(* IEC 61131-3 sources: NachHouse_TST/API/pilot_Api_V11, 8 files *)

(* ---- 07_Nh_JsonRamTest.st ---- *)
// One-shot transport measurement. The records are synthetic because the production mRam is not populated yet.
// Files intentionally remain in //RAM/NACHHOUSE/ for manual inspection after the test.

TYPE
  NH_REC_ALL {PUBLIC}  {HIDDEN}: STRUCT 	// uvodny zaznam pre vsetky DEV alebo struktury, ktore su tabulkou
 	  Ok              : BOOL := TRUE; // platna veta = NOT DELTED
    ID              : INT;					// identifikator zaznamu {Rec Number}
  END_STRUCT;

  NH_CFG_ALL	{PUBLIC}  {HIDDEN}: STRUCT 	// univerzalne CFG pre vsetky DEV
    RoomID          : INT;			    // do ktorej miestnosti patri toto DEV
    CategoryID      : INT;					// domovska kategoria Device
  END_STRUCT;

  NH_JSON_TEST_ROOM  {PUBLIC} : STRUCT    // povodna testovacia struktura
    // povodna testovacia struktura
    RoomId          : UDINT;
    LightLevel      : UINT;
    Temperature10   : INT;
    Online          : BOOL;
   END_STRUCT

  NH_JSON_MEM  {PUBLIC} : STRUCT    // toto zoberiema ako STATE  a bude cele v mRam ako struktura, ktora sa bude posielat do JSON-stat
    rec             : NH_REC_ALL;   // hlavicka - ked sa bude posielat do JSON len stat = mRam
    all             : NH_CFG_ALL;   // premenn, ktore sa pouzivaju casto pri behu programu, ale nemenia sa
    sta             : NH_JSON_TEST_ROOM;   // hlavnme stavove premenne
   END_STRUCT

  NH_JSON_TEST_ROOM_CFG {PUBLIC} : STRUCT   // konfiguracia ulozena
    rec             : NH_REC_ALL;   // duplicitna hlavicka - ked sa bude posielat do JSON len config
    Name            : STRING[32];  // nazov miestnosti
    // iba pre testivanie  STRUCT <-> JSON (ostatnych elementarnych typov, ktore mozu byt STRUCT -> JSON)
    _Dint           : DINT;
    _Sint           : SINT;
    _Usint          : USINT;
    _Uint           : USINT;
    _Real           : REAL;
    _LReal          : LREAL;
    _String         : STRING[30];   // prazdny string
    _StringCZSK     : STRING := 'SVKBEGIN_ščľťžýáíé_SVKEND';   // string obsahujuci ceske a slovenske znaky
    _BYTE           : BYTE;
    _WORD           : WORD;
    _TIME           : TIME;
    _DATE           : DATE;
    _TIME_OF_DAY    : TOD;
    _DATE_AND_TIME  : DT;
   END_STRUCT

  NH_LIGT {PUBLIC}  : STRUCT    // toto je kompletna premenn v nasom pripade JSON, inak NH_ROOM, NH_BLIND,NH_HEAT ...
    mem             : NH_JSON_MEM;             // co budes v mRam ako STATE (memory) - RAM je pouzita na disku '/RAM/'
    cfg             : NH_JSON_TEST_ROOM_CFG;   // toto bude len na SDC
   END_STRUCT

(*
   NH_JSON_TEST_ROOM : STRUCT
      RoomId          : UDINT;
      LightLevel      : UINT;
      Temperature10   : INT;
      Online          : BOOL;
   END_STRUCT
*)
END_TYPE

VAR_GLOBAL CONSTANT
  NH_JSON_TEST_RECORDS : UINT := 300;
  // Historical prototype declaration; unused and not valid in VAR_GLOBAL CONSTANT.
  // aNhJSON {PUBLIC} {TRACK_ADR} {OPEN_UP} : NH_LIGHT;
END_VAR

VAR_GLOBAL
   NhJsonTestRooms        : ARRAY[1..300] OF NH_JSON_TEST_ROOM;
   NhJsonTestInitialized  : BOOL := FALSE;
   NhJsonTestState        : USINT := 0;
   NhJsonTestMode         : USINT := 0;
   NhJsonTestIndex        : UINT := 0;
   NhJsonTestHandle       : HANDLE := INVALID_HANDLE_VALUE;
   NhJsonTestWritten      : UDINT := 0;
   NhJsonTestBuildCycles  : UINT := 0;
   NhJsonTestFileName     : STRING[80];
END_VAR

FUNCTION NhJsonTestWrite : BOOL
   VAR_INPUT
      Text : STRING[255];
   END_VAR
   VAR
      Count : UDINT;
   END_VAR
   NhJsonTestWrite := FALSE;
   Count := FileWrite(hFile := NhJsonTestHandle, adrBuf := PTR_TO_UDINT(ADR(Text)), size := UINT_TO_UDINT(LEN(Text)));
   IF Count <> UINT_TO_UDINT(LEN(Text)) THEN RETURN; END_IF;
   NhJsonTestWritten := NhJsonTestWritten + Count;
   NhJsonTestWrite := TRUE;
END_FUNCTION

FUNCTION NhJsonTestWriteRecord : BOOL
   VAR_INPUT
      Index  : UINT;
      Prefix : BOOL;
   END_VAR
   VAR
      Record : PTR_TO NH_JSON_TEST_ROOM;
      Line   : STRING[255];
      Online : STRING[5];
   END_VAR
   NhJsonTestWriteRecord := FALSE;
   Record := ADR(NhJsonTestRooms[Index]);
   IF Record^.Online THEN Online := 'true'; ELSE Online := 'false'; END_IF;
   IF Prefix THEN Line := ','; ELSE Line := ''; END_IF;
   Line := CONCAT(Line, '{"id":', UDINT_TO_STRING(Record^.RoomId), ',"level":', UINT_TO_STRING(Record^.LightLevel), ',"temperature10":', INT_TO_STRING(Record^.Temperature10), ',"online":', Online, '}');
   NhJsonTestWriteRecord := NhJsonTestWrite(Text := Line);
END_FUNCTION

FUNCTION NhJsonTestInitialize : BOOL
   VAR
      Index : UINT;
   END_VAR
   NhJsonTestInitialize := NhJsonTestInitialized;
   IF NhJsonTestInitialized THEN RETURN; END_IF;
   FOR Index := 1 TO NH_JSON_TEST_RECORDS DO
      NhJsonTestRooms[Index].RoomId := UINT_TO_UDINT(Index);
      NhJsonTestRooms[Index].LightLevel := (Index * 7) MOD 101;
      NhJsonTestRooms[Index].Temperature10 := 185 + UINT_TO_INT(Index MOD 65);
      NhJsonTestRooms[Index].Online := (Index MOD 11) <> 0;
   END_FOR;
   NhJsonTestInitialized := TRUE;
   NhJsonTestInitialize := TRUE;
END_FUNCTION

FUNCTION NhJsonTestCycle : BOOL
   VAR
      Index : UINT;
      Header : STRING[255];
      Trailer : STRING[255];
      ModeText : STRING[6];
      Closed : BOOL;
   END_VAR
   NhJsonTestCycle := FALSE;
   NhJsonTestInitialize();
   IF System_S.LAST_CYCLE_TIME_100US > NhJsonTestMaxCycle100us THEN NhJsonTestMaxCycle100us := System_S.LAST_CYCLE_TIME_100US; END_IF;
   CASE NhJsonTestState OF
      0:
         IF (NhJsonTestCommand = 1) OR (NhJsonTestCommand = 2) THEN
            NhJsonTestMode := NhJsonTestCommand; NhJsonTestCommand := 0; NhJsonTestStatus := NhJsonTestMode;
            NhJsonTestBytes := 0; NhJsonTestRecords := 0; NhJsonTestMaxCycle100us := 0; NhJsonTestWritten := 0; NhJsonTestBuildCycles := 0; NhJsonTestState := 1;
         END_IF;
      1:
         IF NhJsonTestMode = 1 THEN NhJsonTestFileName := '//RAM/NACHHOUSE/nh-json-test-stream.json'; ELSE NhJsonTestFileName := '//RAM/NACHHOUSE/nh-json-test-burst.json'; END_IF;
         NhJsonTestHandle := FileOpen(fileName := NhJsonTestFileName, mode := F_WRITE);
         IF NhJsonTestHandle = INVALID_HANDLE_VALUE THEN NhJsonTestStatus := 255; NhJsonTestState := 0; RETURN; END_IF;
         IF NhJsonTestMode = 1 THEN
            ModeText := 'stream';
         ELSE
            ModeText := 'burst';
         END_IF;
         Header := CONCAT('{"protocol":1,"kind":"patch","sequence":', UDINT_TO_STRING(NhTxRevision + 1), ',"baseSequence":', UDINT_TO_STRING(NhTxRevision), ',"mode":"', ModeText, '","groups":[{"type":"ROOMS","schema":"NH_JSON_TEST_ROOM","records":[');
         IF NOT NhJsonTestWrite(Text := Header) THEN NhJsonTestStatus := 255; NhJsonTestState := 4; RETURN; END_IF;
         NhJsonTestIndex := 1; NhJsonTestState := 2;
      2:
         IF NhJsonTestMode = 1 THEN
            IF NOT NhJsonTestWriteRecord(Index := NhJsonTestIndex, Prefix := NhJsonTestIndex > 1) THEN NhJsonTestStatus := 255; NhJsonTestState := 4; RETURN; END_IF;
            NhJsonTestIndex := NhJsonTestIndex + 1; NhJsonTestBuildCycles := NhJsonTestBuildCycles + 1;
         ELSE
            FOR Index := 1 TO NH_JSON_TEST_RECORDS DO
               IF NOT NhJsonTestWriteRecord(Index := Index, Prefix := Index > 1) THEN NhJsonTestStatus := 255; NhJsonTestState := 4; RETURN; END_IF;
            END_FOR;
            NhJsonTestIndex := NH_JSON_TEST_RECORDS + 1; NhJsonTestBuildCycles := 1;
         END_IF;
         IF NhJsonTestIndex > NH_JSON_TEST_RECORDS THEN NhJsonTestState := 3; END_IF;
      3:
         Trailer := CONCAT(']}],"metrics":{"records":', UINT_TO_STRING(NH_JSON_TEST_RECORDS), ',"buildCycles":', UINT_TO_STRING(NhJsonTestBuildCycles), '}}');
         IF NOT NhJsonTestWrite(Text := Trailer) THEN NhJsonTestStatus := 255; NhJsonTestState := 4; RETURN; END_IF;
         Closed := FileClose(hFile := NhJsonTestHandle); NhJsonTestHandle := INVALID_HANDLE_VALUE;
         IF NOT Closed THEN NhJsonTestStatus := 255; NhJsonTestState := 0; RETURN; END_IF;
         NhJsonTestBytes := NhJsonTestWritten; NhJsonTestRecords := NH_JSON_TEST_RECORDS; NhTxRevision := NhTxRevision + 1; NhJsonTestStatus := 3; NhJsonTestState := 0;
      4:
         IF NhJsonTestHandle <> INVALID_HANDLE_VALUE THEN FileClose(hFile := NhJsonTestHandle); NhJsonTestHandle := INVALID_HANDLE_VALUE; END_IF;
         NhJsonTestState := 0;
   END_CASE;
   NhJsonTestCycle := TRUE;
END_FUNCTION

(* ---- 01_Nh_Api_STRUCT.st ---- *)
// NachHouse API V11: one shared RX mailbox, one shared TX buffer and one transaction owner.
// SK: NachHouse API V11: jeden spolocny RX mailbox, jeden TX buffer a jeden vlastnik transakcie.

VAR_GLOBAL CONSTANT
   NH_API_VERSION                 : UINT := 11;           // Public binary API format version. SK: Verzia verejneho binarneho API formatu.
   NH_API_MAGIC                   : DWORD := 16#5041484E; // ASCII NHAP in little-endian byte order. SK: ASCII NHAP v little-endian poradi bajtov.
   NH_API_HEADER_SIZE             : UINT := 40;           // Fixed frame header size in bytes. SK: Pevna velkost hlavicky ramca v bajtoch.
   NH_API_TX_WORD_COUNT           : UINT := 512;          // Shared TX capacity in DWORD words. SK: Kapacita spolocneho TX pola v DWORD.
   NH_API_RX_WORD_COUNT           : UINT := 64;           // Shared RX capacity in DWORD words. SK: Kapacita spolocneho RX pola v DWORD.
   NH_API_TX_BYTE_CAPACITY        : UINT := 2048;         // Shared TX capacity in bytes. SK: Kapacita spolocneho TX pola v bajtoch.
   NH_API_RX_BYTE_CAPACITY        : UINT := 256;          // Shared RX capacity in bytes. SK: Kapacita spolocneho RX pola v bajtoch.
   NH_API_MAX_ROOMS               : UINT := 40;           // Maximum number of pilot room records. SK: Najvacsi pocet room zaznamov pilotu.
   NH_LOAD_DEVICE_COUNT           : UINT := 800;          // Number of compact smart-home model devices. SK: Pocet kompaktnych modelovych smart-home zariadeni.
   NH_API_TRANSACTION_TIMEOUT_MS  : UDINT := 30000;       // Maximum owner inactivity time. SK: Maximalny cas necinnosti vlastnika.
   NH_API_BROADCAST_HOLD_MS       : UDINT := 500;         // Minimum time one best-effort broadcast frame stays stable. SK: Minimalny cas stability jedneho broadcast ramca.

   NH_API_CONFIG_RECORD_SIZE      : UINT := 138;          // Wire size of one room config record. SK: Wire velkost jedneho room config zaznamu.
   NH_API_STATE_RECORD_SIZE       : UINT := 22;           // Wire size of one room state record. SK: Wire velkost jedneho room state zaznamu.
   NH_API_CONFIG_DIFF_SIZE        : UINT := 143;          // Operation, RoomId and config record. SK: Operacia, RoomId a config zaznam.
   NH_API_STATE_DIFF_SIZE         : UINT := 27;           // Operation, RoomId and state record. SK: Operacia, RoomId a state zaznam.
   NH_API_CONFIG_PER_FRAME        : USINT := 14;           // Config records fitting into one TX frame. SK: Config zaznamy, ktore sa zmestia do jedneho TX ramca.
   NH_API_STATE_PER_FRAME         : USINT := 40;           // State records fitting into one TX frame. SK: State zaznamy, ktore sa zmestia do jedneho TX ramca.
   NH_API_CONFIG_DIFF_PER_FRAME   : USINT := 14;           // Config changes fitting into one TX frame. SK: Config zmeny, ktore sa zmestia do jedneho TX ramca.
   NH_API_STATE_DIFF_PER_FRAME    : USINT := 40;           // State changes fitting into one TX frame. SK: State zmeny, ktore sa zmestia do jedneho TX ramca.

   NH_API_STATE_IDLE              : UINT := 0;             // No transaction owns the API. SK: API nevlastni ziadna transakcia.
   NH_API_STATE_OWNER_READY       : UINT := 1;             // PLC accepted OwnerClientId; owner may write RX. SK: PLC prijalo OwnerClientId; vlastnik moze zapisat RX.
   NH_API_STATE_RX_READY          : UINT := 2;             // Owner completed RX and committed it. SK: Vlastnik dokoncil RX a potvrdil ho.

   NH_API_MODE_NONE               : USINT := 0;            // No frame sequence is active. SK: Nie je aktivna ziadna sekvencia ramcov.
   NH_API_MODE_SNAPSHOT           : USINT := 1;            // Targeted snapshot sequence. SK: Cielena snapshot sekvencia.
   NH_API_MODE_COMMAND            : USINT := 2;            // Targeted command response sequence. SK: Cielena sekvencia odpovede na prikaz.
   NH_API_MODE_BROADCAST_DIFF     : USINT := 3;            // Best-effort PLC-originated diff. SK: Best-effort diff vyvolany PLC.
   NH_API_MODE_BROADCAST_SNAPSHOT : USINT := 4;            // Best-effort test snapshot without an owner. SK: Best-effort test snapshot bez vlastnika.

   NH_API_MSG_SNAPSHOT_REQUEST    : UINT := 1;             // RX request for current room snapshot. SK: RX poziadavka na aktualny room snapshot.
   NH_API_MSG_ADD_ROOM            : UINT := 2;             // RX request to add a room. SK: RX poziadavka na pridanie miestnosti.
   NH_API_MSG_DELETE_ROOM         : UINT := 3;             // RX request to delete a room. SK: RX poziadavka na zmazanie miestnosti.
   NH_API_MSG_COPY_ROOM           : UINT := 4;             // RX request to copy a room. SK: RX poziadavka na kopirovanie miestnosti.
   NH_API_MSG_SET_ROOM_CONFIG     : UINT := 5;             // RX request to replace room config. SK: RX poziadavka na nahradenie room configu.
   NH_API_MSG_SET_ROOM_STATE      : UINT := 6;             // RX request to replace room state. SK: RX poziadavka na nahradenie room state.
   NH_API_MSG_CONFIG_SNAPSHOT     : UINT := 101;           // TX config snapshot part. SK: TX cast config snapshotu.
   NH_API_MSG_STATE_SNAPSHOT      : UINT := 102;           // TX state snapshot part. SK: TX cast state snapshotu.
   NH_API_MSG_CONFIG_DIFF         : UINT := 103;           // TX config changes. SK: TX zmeny configu.
   NH_API_MSG_STATE_DIFF          : UINT := 104;           // TX state changes. SK: TX zmeny state.
   NH_API_MSG_SNAPSHOT_DONE       : UINT := 105;           // TX final snapshot frame. SK: TX posledny ramec snapshotu.
   NH_API_MSG_RESULT              : UINT := 106;           // TX final command result. SK: TX konecny vysledok prikazu.

   NH_API_SCHEMA_NONE             : UINT := 0;             // Frame has no structured record. SK: Ramec nema strukturovany zaznam.
   NH_API_SCHEMA_ROOM_CONFIG      : UINT := 1;             // NH_ROOM_CONFIG wire schema. SK: Wire schema NH_ROOM_CONFIG.
   NH_API_SCHEMA_ROOM_STATE       : UINT := 2;             // NH_ROOM_STATE wire schema. SK: Wire schema NH_ROOM_STATE.

   NH_API_CHANGE_UPSERT           : USINT := 1;            // Add or complete record replacement. SK: Pridanie alebo uplne nahradenie zaznamu.
   NH_API_CHANGE_DELETE           : USINT := 2;            // Record deletion. SK: Zmazanie zaznamu.

   NH_API_RESULT_NONE             : USINT := 0;            // No result is available. SK: Vysledok nie je k dispozicii.
   NH_API_RESULT_OK               : USINT := 1;            // Request completed successfully. SK: Poziadavka bola uspesna.
   NH_API_RESULT_BUSY             : USINT := 2;            // API is owned by another transaction. SK: API vlastni ina transakcia.
   NH_API_RESULT_BAD_FRAME        : USINT := 3;            // Header, size, owner or CRC is invalid. SK: Hlavicka, velkost, vlastnik alebo CRC su neplatne.
   NH_API_RESULT_NOT_FOUND        : USINT := 4;            // Requested room does not exist. SK: Pozadovana miestnost neexistuje.
   NH_API_RESULT_NO_FREE_SLOT     : USINT := 5;            // No internal room slot is free. SK: Nie je volny interny room slot.
   NH_API_RESULT_ALREADY_EXISTS   : USINT := 6;            // Target RoomId already exists. SK: Cielove RoomId uz existuje.
   NH_API_RESULT_INVALID          : USINT := 7;            // Request payload is invalid. SK: Payload poziadavky nie je platny.
   NH_API_RESULT_UNSUPPORTED      : USINT := 8;            // Message type is unsupported. SK: Typ spravy nie je podporovany.
   NH_API_RESULT_TIMEOUT          : USINT := 9;            // Owner did not complete the handshake. SK: Vlastnik nedokoncil handshake.

   NH_API_TEST_NONE               : USINT := 0;            // Test interface performs no action. SK: Testovacie rozhranie nevykona akciu.
   NH_API_TEST_SET_STATE          : USINT := 1;            // Test interface changes room state. SK: Testovacie rozhranie zmeni room state.
   NH_API_TEST_ADD_ROOM           : USINT := 2;            // Test interface adds a room. SK: Testovacie rozhranie prida miestnost.
   NH_API_TEST_DELETE_ROOM        : USINT := 3;            // Test interface deletes a room. SK: Testovacie rozhranie zmaze miestnost.
   NH_API_TEST_COPY_ROOM          : USINT := 4;            // Test interface copies a room. SK: Testovacie rozhranie skopiruje miestnost.
   NH_API_TEST_SET_CONFIG         : USINT := 5;            // Test interface changes room config. SK: Testovacie rozhranie zmeni room config.
   NH_API_TEST_REQUEST_SNAPSHOT   : USINT := 6;            // Test interface publishes a broadcast snapshot. SK: Testovacie rozhranie publikuje broadcast snapshot.
   NH_API_TEST_AWAY               : USINT := 7;            // Test interface applies the LOAD_800 departure scene. SK: Testovacie rozhranie vykona modelovu scenu odchod LOAD_800.
END_VAR

TYPE
   NH_ROOM_CONFIG : STRUCT // Static room configuration used by snapshots, diffs and commands. SK: Staticka konfiguracia miestnosti pouzita v snapshotoch, diffoch a prikazoch.
      Used           : BOOL;       // TRUE marks an occupied internal slot. SK: TRUE oznacuje obsadeny interny slot.
      RoomId         : UDINT;      // Stable room identifier. SK: Stabilny identifikator miestnosti.
      Name           : STRING[64]; // UTF-8 room name, at most 64 bytes. SK: UTF-8 nazov miestnosti, najviac 64 bajtov.
      ProjectName    : STRING[64]; // UTF-8 project name, at most 64 bytes. SK: UTF-8 projektovy nazov, najviac 64 bajtov.
      IconId         : UINT;       // Client icon identifier. SK: Identifikator ikony klienta.
      SortDefault    : UINT;       // Default room order. SK: Predvolene poradie miestnosti.
   END_STRUCT

   NH_ROOM_STATE : STRUCT // Dynamic room state used by snapshots, diffs and commands. SK: Dynamicky stav miestnosti pouzity v snapshotoch, diffoch a prikazoch.
      RoomId         : UDINT;      // Stable ID matching the config record. SK: Stabilne ID zodpovedajuce config zaznamu.
      Temperature    : REAL;       // Temperature in degrees Celsius. SK: Teplota v stupnoch Celzia.
      Humidity       : REAL;       // Relative humidity in percent. SK: Relativna vlhkost v percentach.
      Presence       : BOOL;       // Presence flag. SK: Priznak pritomnosti.
      DayPhase       : UINT;       // Day-phase icon identifier. SK: Identifikator ikony fazy dna.
      CategoryMask   : DWORD;      // Bit mask of active categories. SK: Bitova maska aktivnych kategorii.
      AlarmLevel     : USINT;      // Alarm level from 0 to 2. SK: Uroven alarmu od 0 do 2.
      Online         : BOOL;       // Room data availability. SK: Dostupnost dat miestnosti.
      Twilight       : BOOL;       // Twilight state used by room browser. SK: Stav osvetlenia pouzity room browserom.
   END_STRUCT

   NH_API_INFO : STRUCT // Minimal global owner and handshake state. SK: Minimalny globalny stav vlastnika a handshake.
      ApiVersion      : UINT;      // Binary API contract version. SK: Verzia binarneho API kontraktu.
      State           : UINT;      // Zero is free; nonzero is the current handshake step. SK: Nula je volno; nenulova hodnota je aktualny handshake krok.
      OwnerClientId   : UDINT;     // Fresh nonzero owner token of the current transaction. SK: Novy nenulovy token vlastnika aktualnej transakcie.
   END_STRUCT

   NH_API_TEST_CONTROL : STRUCT // Direct WebMaker/debug interface for PLC-originated test changes. SK: Priame WebMaker/debug rozhranie pre testovacie zmeny vyvolane PLC.
      Execute         : BOOL;       // Set TRUE last to execute the prepared action. SK: Nastavit TRUE ako posledne pre vykonanie pripravenej akcie.
      Finished        : BOOL;       // TRUE after the test action was accepted. SK: TRUE po prijati testovacej akcie.
      Action          : USINT;      // Requested NH_API_TEST_* action. SK: Pozadovana akcia NH_API_TEST_*.
      ResultCode      : USINT;      // NH_API_RESULT_* outcome. SK: Vysledok NH_API_RESULT_*.
      RoomId          : UDINT;      // Target room ID. SK: Cielove ID miestnosti.
      SourceRoomId    : UDINT;      // Source ID for copy. SK: Zdrojove ID pri kopirovani.
      Name            : STRING[64]; // New room name. SK: Novy nazov miestnosti.
      ProjectName     : STRING[64]; // New project name. SK: Novy projektovy nazov.
      IconId          : UINT;       // New icon identifier. SK: Novy identifikator ikony.
      Temperature     : REAL;       // Test temperature. SK: Testovacia teplota.
      Humidity        : REAL;       // Test humidity. SK: Testovacia vlhkost.
      Presence        : BOOL;       // Test presence. SK: Testovacia pritomnost.
      DayPhase        : UINT;       // Test day phase. SK: Testovacia faza dna.
      CategoryMask    : DWORD;      // Test category mask. SK: Testovacia maska kategorii.
      AlarmLevel      : USINT;      // Test alarm level. SK: Testovacia uroven alarmu.
      Online          : BOOL;       // Test availability. SK: Testovacia dostupnost.
      Twilight        : BOOL;       // Test twilight state. SK: Testovaci twilight stav.
   END_STRUCT

   NH_LOAD_TEST_STATUS : STRUCT // Observable LOAD_800 test status. SK: Pozorovatelny stav testu LOAD_800.
      DepartureActive : BOOL;  // TRUE while the model is in departure mode. SK: TRUE pocas modeloveho rezimu odchod.
      LastChangedCount: UINT;  // Device records changed by the last scene. SK: Pocet zaznamov zmenenych poslednou scenou.
      LastApplyMs     : UDINT; // PLC time spent applying the scene. SK: Cas PLC potrebny na vykonanie sceny.
      Sequence        : UDINT; // Increments after every completed model scene. SK: Zvysi sa po kazdej dokoncenej modelovej scene.
   END_STRUCT
END_TYPE

VAR_GLOBAL
   NhApiInfo       {PUBLIC_API} : NH_API_INFO;                // Minimal global transaction control. SK: Minimalne globalne riadenie transakcie.
   NhApiTX                      : ARRAY[0..511] OF DWORD;     // Internal frame published as one binary WWW file. SK: Interny ramec publikovany ako jeden binarny WWW subor.
   NhApiRX                      : ARRAY[0..63] OF DWORD;      // Internal owner-to-PLC request frame decoded from Base64 transport.
   NhApiTest       {PUBLIC_API} : NH_API_TEST_CONTROL;        // Direct PLC-originated test control. SK: Priame riadenie testov vyvolanych PLC.
   NhLoadTest      {PUBLIC_API} : NH_LOAD_TEST_STATUS;        // LOAD_800 status and measurements. SK: Stav a merania LOAD_800.
   NhLoadDevices                : ARRAY[1..800] OF DWORD;     // Internal load-test model; never publish array elements through PLCComS diffs.

   // JSON RAM transport test: only NhTxRevision is the client-ready signal.
   NhTxRevision     {PUBLIC_API} : UDINT := 0;
   NhJsonTestCommand{PUBLIC_API} : USINT := 0; // 1=stream one record/cycle, 2=burst all records/one cycle.
   NhJsonTestStatus {PUBLIC_API} : USINT := 0; // 0=idle, 1=streaming, 2=bursting, 3=ready, 255=error.
   NhJsonTestBytes  {PUBLIC_API} : UDINT := 0;
   NhJsonTestRecords{PUBLIC_API} : UINT := 0;
   NhJsonTestMaxCycle100us {PUBLIC_API} : UINT := 0;

   NhRoomsConfig                : ARRAY[1..40] OF NH_ROOM_CONFIG; // Authoritative PLC room configuration. SK: Autoritativna PLC konfiguracia miestnosti.
   NhRoomsState                 : ARRAY[1..40] OF NH_ROOM_STATE;  // Authoritative PLC room state. SK: Autoritativny PLC stav miestnosti.
END_VAR

VAR_GLOBAL
   NhApiInitialized             : BOOL;                         // One-time initialization completed. SK: Jednorazova inicializacia dokoncena.
   NhActiveOwnerClientId        : UDINT;                        // Owner token captured by PLC. SK: Token vlastnika zachyteny PLC.
   NhExpectedState              : UINT;                         // State value currently owned by PLC. SK: Hodnota State aktualne vlastnena PLC.
   NhTransactionMode           : USINT;                        // Active NH_API_MODE_*. SK: Aktivny NH_API_MODE_*.
   NhTransactionLastMs         : UDINT;                        // Time of the last accepted handshake step. SK: Cas posledneho prijateho handshake kroku.
   NhPublishedFrameId          : UDINT;                        // Monotonic identity of every published TX frame. SK: Monotonny identifikator kazdeho publikovaneho TX ramca.
   NhCommandResult             : USINT;                        // Result sent in the final command frame. SK: Vysledok poslany v poslednom prikazovom ramci.
   NhResultPending             : BOOL;                         // Final command result still has to be sent. SK: Konecny vysledok prikazu este treba odoslat.

   NhConfigShadow              : ARRAY[1..40] OF NH_ROOM_CONFIG; // Last published config image. SK: Posledny publikovany obraz konfiguracie.
   NhStateShadow               : ARRAY[1..40] OF NH_ROOM_STATE;  // Last published state image. SK: Posledny publikovany obraz stavu.

   NhPendingConfig             : ARRAY[1..40] OF NH_ROOM_CONFIG; // Frozen config diff records. SK: Zmrazene zaznamy config diffu.
   NhPendingConfigOperation    : ARRAY[1..40] OF USINT;          // Operations of config diff records. SK: Operacie zaznamov config diffu.
   NhPendingConfigRoomId       : ARRAY[1..40] OF UDINT;          // Stable IDs of config changes. SK: Stabilne ID config zmien.
   NhPendingConfigCount        : USINT;                          // Number of frozen config changes. SK: Pocet zmrazenych config zmien.
   NhPendingConfigNext         : USINT;                          // First config change in the next frame. SK: Prva config zmena v dalsom ramci.
   NhPendingConfigPart         : USINT;                          // Next config diff part index. SK: Index dalsej casti config diffu.
   NhPendingConfigParts        : USINT;                          // Total config diff part count. SK: Celkovy pocet casti config diffu.

   NhPendingState              : ARRAY[1..40] OF NH_ROOM_STATE;  // Frozen state diff records. SK: Zmrazene zaznamy state diffu.
   NhPendingStateOperation     : ARRAY[1..40] OF USINT;          // Operations of state diff records. SK: Operacie zaznamov state diffu.
   NhPendingStateRoomId        : ARRAY[1..40] OF UDINT;          // Stable IDs of state changes. SK: Stabilne ID state zmien.
   NhPendingStateCount         : USINT;                          // Number of frozen state changes. SK: Pocet zmrazenych state zmien.
   NhPendingStateNext          : USINT;                          // First state change in the next frame. SK: Prva state zmena v dalsom ramci.
   NhPendingStatePart          : USINT;                          // Next state diff part index. SK: Index dalsej casti state diffu.
   NhPendingStateParts         : USINT;                          // Total state diff part count. SK: Celkovy pocet casti state diffu.

   NhSnapshotActive            : BOOL;                           // Frozen snapshot sequence is active. SK: Zmrazena snapshot sekvencia je aktivna.
   NhSnapshotStage             : USINT;                          // 1 config, 2 state, 3 done. SK: 1 config, 2 state, 3 done.
   NhSnapshotNext              : USINT;                          // First snapshot record in the next frame. SK: Prvy snapshot zaznam v dalsom ramci.
   NhSnapshotPart              : USINT;                          // Next snapshot part index. SK: Index dalsej casti snapshotu.
   NhSnapshotParts             : USINT;                          // Part count of the current snapshot section. SK: Pocet casti aktualnej sekcie.
   NhSnapshotCount             : USINT;                          // Number of valid frozen rooms. SK: Pocet platnych miestnosti.
   NhSnapshotConfig            : ARRAY[1..40] OF NH_ROOM_CONFIG; // Frozen config snapshot. SK: Zmrazeny obraz konfiguracie.
   NhSnapshotState             : ARRAY[1..40] OF NH_ROOM_STATE;  // Frozen state snapshot. SK: Zmrazeny obraz stavu.
END_VAR

(* ---- 05_Nh_FileTransport.st ---- *)
// Browser-direct binary transport: PLC writes each complete NHAP frame into the inactive RAM-disk slot.
// Browser receives only NhFileFrameId over WSS and downloads one immutable binary response over HTTPS at /RAM/NACHHOUSE/.

VAR_GLOBAL
   NhFileFrameId    {PUBLIC_API} : UDINT := 0; // Commit written only after FileWrite and FileClose succeed.
   NhFileStatus     {PUBLIC_API} : USINT := 0; // 0 idle/OK, 2 open error, 3 short write, 4 close error, 5 invalid frame.
   NhFileLastBytes  {PUBLIC_API} : UINT := 0;  // Diagnostic only; authoritative length is inside the NHAP header.
   NhFileCycleCount {PUBLIC_API} : UDINT := 0; // Diagnostic proof that the publisher runs in every PLC cycle.

   NhFileInitialized            : BOOL := FALSE;
   NhFileLastPublished          : UDINT := 0;
   NhFileName                   : STRING[80];
   NhFileDirectory              : STRING[80] := '//RAM/NACHHOUSE/';
   NhFileHandle                 : HANDLE := INVALID_HANDLE_VALUE;
   NhFileWritten                : UDINT := 0;
   NhFileClosed                 : BOOL := FALSE;
END_VAR

FUNCTION NhFileTransportCycle : BOOL
   VAR_TEMP
      FrameLength : UINT;
   END_VAR

   NhFileTransportCycle := FALSE;
   NhFileCycleCount := NhFileCycleCount + 1;

   IF NOT NhFileInitialized THEN
      // DirCreate may return FALSE when the directory already exists; opening the file is the decisive check.
      DirCreate(dirName := NhFileDirectory);
      NhFileInitialized := TRUE;
   END_IF;

   IF (NhPublishedFrameId = 0) OR (NhPublishedFrameId = NhFileLastPublished) THEN
      NhFileTransportCycle := TRUE;
      RETURN;
   END_IF;

   FrameLength := UDINT_TO_UINT(NhApiReadU32(Buffer := ADR(NhApiTX), Offset := 28));
   IF (FrameLength < NH_API_HEADER_SIZE) OR (FrameLength > NH_API_TX_BYTE_CAPACITY) THEN
      NhFileStatus := 5;
      RETURN;
   END_IF;

   IF (NhPublishedFrameId MOD 2) = 0 THEN
      NhFileName := '//RAM/NACHHOUSE/nhapi-0.bin';
   ELSE
      NhFileName := '//RAM/NACHHOUSE/nhapi-1.bin';
   END_IF;

   NhFileHandle := FileOpen(fileName := NhFileName, mode := F_WRITE);
   IF NhFileHandle = INVALID_HANDLE_VALUE THEN
      NhFileStatus := 2;
      RETURN;
   END_IF;

   NhFileWritten := FileWrite(hFile := NhFileHandle, adrBuf := PTR_TO_UDINT(ADR(NhApiTX)), size := UINT_TO_UDINT(FrameLength));
   NhFileClosed := FileClose(hFile := NhFileHandle);
   NhFileHandle := INVALID_HANDLE_VALUE;

   IF NhFileWritten <> UINT_TO_UDINT(FrameLength) THEN
      NhFileStatus := 3;
      RETURN;
   END_IF;
   IF NOT NhFileClosed THEN
      NhFileStatus := 4;
      RETURN;
   END_IF;

   NhFileLastBytes := FrameLength;
   NhFileStatus := 0;
   NhFileLastPublished := NhPublishedFrameId;
   NhFileFrameId := NhPublishedFrameId; // Application-level commit: always publish last.
   NhFileTransportCycle := TRUE;
END_FUNCTION

(* ---- 06_Nh_RxTextTransport.st ---- *)
// Legacy RX prototype. PLCComS STRING-length capability is verified separately.

VAR_GLOBAL
   NhRxText        {PUBLIC_API} : ARRAY[0..4] OF STRING[80];
   NhRxTextCommit  {PUBLIC_API} : UDINT := 0;
   NhRxTextStatus  {PUBLIC_API} : USINT := 0; // 0 idle/OK, 1 invalid Base64, 2 invalid decoded length.
   NhRxTextBytes   {PUBLIC_API} : UINT := 0;
   NhRxLastCommit               : UDINT := 0;
END_VAR

FUNCTION NhBase64Value : INT
   VAR_INPUT
      Character : BYTE;
   END_VAR
   IF (Character >= 65) AND (Character <= 90) THEN
      NhBase64Value := BYTE_TO_INT(Character) - 65;
   ELSIF (Character >= 97) AND (Character <= 122) THEN
      NhBase64Value := BYTE_TO_INT(Character) - 71;
   ELSIF (Character >= 48) AND (Character <= 57) THEN
      NhBase64Value := BYTE_TO_INT(Character) + 4;
   ELSIF Character = 43 THEN
      NhBase64Value := 62;
   ELSIF Character = 47 THEN
      NhBase64Value := 63;
   ELSIF Character = 61 THEN
      NhBase64Value := -2; // '=' padding
   ELSE
      NhBase64Value := -1;
   END_IF;
END_FUNCTION

FUNCTION NhDecodeBase64Chunk : INT
   VAR_INPUT
      Text       : STRING[80];
      DestOffset : UINT;
   END_VAR
   VAR
      Source     : PTR_TO BYTE;
      Target     : PTR_TO BYTE;
      TextLength : UINT;
      Index      : UINT;
      Written    : UINT;
      V0         : INT;
      V1         : INT;
      V2         : INT;
      V3         : INT;
   END_VAR

   NhDecodeBase64Chunk := -1;
   TextLength := INT_TO_UINT(LEN(Text));
   IF TextLength = 0 THEN NhDecodeBase64Chunk := 0; RETURN; END_IF;
   IF (TextLength MOD 4) <> 0 THEN RETURN; END_IF;
   Source := ADR(Text);
   Target := ADR(NhApiRX) + UINT_TO_UDINT(DestOffset);
   Index := 0;
   Written := 0;

   WHILE Index < TextLength DO
      V0 := NhBase64Value(Character := Source^); Source := Source + 1;
      V1 := NhBase64Value(Character := Source^); Source := Source + 1;
      V2 := NhBase64Value(Character := Source^); Source := Source + 1;
      V3 := NhBase64Value(Character := Source^); Source := Source + 1;
      IF (V0 < 0) OR (V1 < 0) OR (V2 = -1) OR (V3 = -1) THEN RETURN; END_IF;
      IF (DestOffset + Written) >= NH_API_RX_BYTE_CAPACITY THEN RETURN; END_IF;
      Target^ := INT_TO_BYTE((V0 * 4) + (V1 / 16)); Target := Target + 1; Written := Written + 1;
      IF V2 >= 0 THEN
         IF (DestOffset + Written) >= NH_API_RX_BYTE_CAPACITY THEN RETURN; END_IF;
         Target^ := INT_TO_BYTE(((V1 MOD 16) * 16) + (V2 / 4)); Target := Target + 1; Written := Written + 1;
         IF V3 >= 0 THEN
            IF (DestOffset + Written) >= NH_API_RX_BYTE_CAPACITY THEN RETURN; END_IF;
            Target^ := INT_TO_BYTE(((V2 MOD 4) * 64) + V3); Target := Target + 1; Written := Written + 1;
         ELSIF Index + 4 <> TextLength THEN RETURN;
         END_IF;
      ELSIF (V3 <> -2) OR (Index + 4 <> TextLength) THEN RETURN;
      END_IF;
      Index := Index + 4;
   END_WHILE;
   NhDecodeBase64Chunk := UINT_TO_INT(Written);
END_FUNCTION

FUNCTION NhRxTextTransportCycle : BOOL
   VAR
      ChunkIndex : UINT;
      Decoded     : INT;
      Total       : UINT;
      FrameLength : UDINT;
   END_VAR

   NhRxTextTransportCycle := TRUE;
   IF (NhApiInfo.State <> NH_API_STATE_OWNER_READY) OR
      (NhRxTextCommit = 0) OR
      (NhRxTextCommit <> NhApiInfo.OwnerClientId) OR
      (NhRxTextCommit = NhRxLastCommit) THEN RETURN;
   END_IF;

   NhApiClearBuffer(Buffer := ADR(NhApiRX), Length := NH_API_RX_BYTE_CAPACITY);
   Total := 0;
   FOR ChunkIndex := 0 TO 4 DO
      Decoded := NhDecodeBase64Chunk(Text := NhRxText[ChunkIndex], DestOffset := Total);
      IF Decoded < 0 THEN NhRxTextStatus := 1; RETURN; END_IF;
      Total := Total + INT_TO_UINT(Decoded);
   END_FOR;

   IF Total < NH_API_HEADER_SIZE THEN NhRxTextStatus := 2; RETURN; END_IF;
   FrameLength := NhApiReadU32(Buffer := ADR(NhApiRX), Offset := 28);
   IF (FrameLength <> UINT_TO_UDINT(Total)) OR (FrameLength > UINT_TO_UDINT(NH_API_RX_BYTE_CAPACITY)) THEN
      NhRxTextStatus := 2;
      RETURN;
   END_IF;

   NhRxTextBytes := Total;
   NhRxTextStatus := 0;
   NhRxLastCommit := NhRxTextCommit;
   NhApiInfo.State := NH_API_STATE_RX_READY;
END_FUNCTION

(* ---- 02_Nh_Api_UTILS.st ---- *)
// Wire-format helpers have no hidden state. SK: Pomocne funkcie wire formatu su bez skryteho stavu.

FUNCTION NhApiSystemTimeMs : UDINT
   // Returns the PLC system time in milliseconds. SK: Vrati systemovy cas PLC v milisekundach.
   VAR_EXTERNAL
      AT %SL52 : DWORD; // Absolute PLC system-time register. SK: Absolutny systemovy register casu PLC.
   END_VAR
   NhApiSystemTimeMs := DWORD_TO_UDINT(%SL52);
END_FUNCTION

FUNCTION NhApiWriteByte : BOOL
   // Writes one byte at the specified buffer offset. SK: Zapise jeden bajt na zadany offset buffera.
   VAR_INPUT
      Buffer : PTR_TO BYTE; // Start of the destination buffer. SK: Zaciatok cieloveho buffera.
      Offset : UINT;        // Zero-based byte offset. SK: Nulovy byte offset.
      Value  : BYTE;        // Value to write. SK: Zapisovana hodnota.
   END_VAR
   VAR
      Position : PTR_TO BYTE; // Pointer advanced to the target byte. SK: Pointer posunuty na cielovy bajt.
   END_VAR
   Position := Buffer + UINT_TO_UDINT(Offset);
   Position^ := Value;
   NhApiWriteByte := TRUE;
END_FUNCTION

FUNCTION NhApiReadByte : BYTE
   // Reads one byte from the specified buffer offset. SK: Precita jeden bajt zo zadaneho offsetu buffera.
   VAR_INPUT
      Buffer : PTR_TO BYTE; // Start of the source buffer. SK: Zaciatok zdrojoveho buffera.
      Offset : UINT;        // Zero-based byte offset. SK: Nulovy byte offset.
   END_VAR
   VAR
      Position : PTR_TO BYTE; // Pointer advanced to the source byte. SK: Pointer posunuty na zdrojovy bajt.
   END_VAR
   Position := Buffer + UINT_TO_UDINT(Offset);
   NhApiReadByte := Position^;
END_FUNCTION

FUNCTION NhApiWriteU16 : BOOL
   // Writes a 16-bit value in little-endian format. SK: Zapise 16-bitovu hodnotu vo formate little-endian.
   VAR_INPUT
      Buffer : PTR_TO BYTE; // Destination byte buffer. SK: Cielovy byte buffer.
      Offset : UINT;        // Zero-based byte offset. SK: Nulovy byte offset.
      Value  : UINT;        // Value written little-endian. SK: Hodnota zapisovana little-endian.
   END_VAR
   NhApiWriteByte(Buffer := Buffer, Offset := Offset, Value := WORD_TO_BYTE(UINT_TO_WORD(Value) AND 16#00FF));
   NhApiWriteByte(Buffer := Buffer, Offset := Offset + 1, Value := WORD_TO_BYTE(SHR(UINT_TO_WORD(Value), 8)));
   NhApiWriteU16 := TRUE;
END_FUNCTION

FUNCTION NhApiWriteU32 : BOOL
   // Writes a 32-bit value in little-endian format. SK: Zapise 32-bitovu hodnotu vo formate little-endian.
   VAR_INPUT
      Buffer : PTR_TO BYTE; // Destination byte buffer. SK: Cielovy byte buffer.
      Offset : UINT;        // Zero-based byte offset. SK: Nulovy byte offset.
      Value  : UDINT;       // Value written little-endian. SK: Hodnota zapisovana little-endian.
   END_VAR
   VAR
      Raw : DWORD;          // Bit image of the value. SK: Bitovy obraz hodnoty.
   END_VAR
   Raw := UDINT_TO_DWORD(Value);
   NhApiWriteByte(Buffer := Buffer, Offset := Offset, Value := DWORD_TO_BYTE(Raw AND 16#000000FF));
   NhApiWriteByte(Buffer := Buffer, Offset := Offset + 1, Value := DWORD_TO_BYTE(SHR(Raw, 8) AND 16#000000FF));
   NhApiWriteByte(Buffer := Buffer, Offset := Offset + 2, Value := DWORD_TO_BYTE(SHR(Raw, 16) AND 16#000000FF));
   NhApiWriteByte(Buffer := Buffer, Offset := Offset + 3, Value := DWORD_TO_BYTE(SHR(Raw, 24) AND 16#000000FF));
   NhApiWriteU32 := TRUE;
END_FUNCTION

FUNCTION NhApiReadU16 : UINT
   // Reads a 16-bit value in little-endian format. SK: Precita 16-bitovu hodnotu vo formate little-endian.
   VAR_INPUT
      Buffer : PTR_TO BYTE; // Source byte buffer. SK: Zdrojovy byte buffer.
      Offset : UINT;        // Zero-based byte offset. SK: Nulovy byte offset.
   END_VAR
   NhApiReadU16 := WORD_TO_UINT(BYTE_TO_WORD(NhApiReadByte(Buffer := Buffer, Offset := Offset)) OR
      SHL(BYTE_TO_WORD(NhApiReadByte(Buffer := Buffer, Offset := Offset + 1)), 8));
END_FUNCTION

FUNCTION NhApiReadU32 : UDINT
   // Reads a 32-bit value in little-endian format. SK: Precita 32-bitovu hodnotu vo formate little-endian.
   VAR_INPUT
      Buffer : PTR_TO BYTE; // Source byte buffer. SK: Zdrojovy byte buffer.
      Offset : UINT;        // Zero-based byte offset. SK: Nulovy byte offset.
   END_VAR
   VAR
      Raw : DWORD;          // Reassembled little-endian value. SK: Zlozena little-endian hodnota.
   END_VAR
   Raw := BYTE_TO_DWORD(NhApiReadByte(Buffer := Buffer, Offset := Offset));
   Raw := Raw OR SHL(BYTE_TO_DWORD(NhApiReadByte(Buffer := Buffer, Offset := Offset + 1)), 8);
   Raw := Raw OR SHL(BYTE_TO_DWORD(NhApiReadByte(Buffer := Buffer, Offset := Offset + 2)), 16);
   Raw := Raw OR SHL(BYTE_TO_DWORD(NhApiReadByte(Buffer := Buffer, Offset := Offset + 3)), 24);
   NhApiReadU32 := DWORD_TO_UDINT(Raw);
END_FUNCTION

FUNCTION NhApiWriteReal : BOOL
   // Writes a REAL using its 32-bit image. SK: Zapise REAL pomocou jeho 32-bitoveho obrazu.
   VAR_INPUT
      Buffer : PTR_TO BYTE; // Destination byte buffer. SK: Cielovy byte buffer.
      Offset : UINT;        // Zero-based byte offset. SK: Nulovy byte offset.
      Value  : REAL;        // IEC REAL written by bit image. SK: IEC REAL zapisany bitovo.
   END_VAR
   VAR
      RawPtr : PTR_TO DWORD;// Pointer to the REAL bit image. SK: Pointer na bitovy obraz REAL.
   END_VAR
   RawPtr := ADR(Value);
   NhApiWriteU32(Buffer := Buffer, Offset := Offset, Value := DWORD_TO_UDINT(RawPtr^));
   NhApiWriteReal := TRUE;
END_FUNCTION

FUNCTION NhApiReadReal : REAL
   // Reads a REAL from its 32-bit image. SK: Precita REAL z jeho 32-bitoveho obrazu.
   VAR_INPUT
      Buffer : PTR_TO BYTE; // Source byte buffer. SK: Zdrojovy byte buffer.
      Offset : UINT;        // Zero-based byte offset. SK: Nulovy byte offset.
   END_VAR
   VAR
      ResultPtr : PTR_TO DWORD; // Pointer to the result bit image. SK: Pointer na bitovy obraz vysledku.
   END_VAR
   ResultPtr := ADR(NhApiReadReal);
   ResultPtr^ := UDINT_TO_DWORD(NhApiReadU32(Buffer := Buffer, Offset := Offset));
END_FUNCTION

FUNCTION NhApiFrameCrc32 : DWORD
   // Calculates CRC32 while treating header bytes 36..39 as zero. SK: Vypocita CRC32, pricom bajty hlavicky 36..39 povazuje za nuly.
   VAR_INPUT
      Buffer : PTR_TO BYTE; // Start of the complete frame. SK: Zaciatok celeho ramca.
      Length : UINT;        // Header plus payload size. SK: Velkost hlavicky a payloadu.
   END_VAR
   VAR
      Crc       : DWORD;    // Running CRC32 value. SK: Priebezna CRC32 hodnota.
      Current   : BYTE;     // Current byte or zero inside CRC field. SK: Aktualny bajt alebo nula v CRC poli.
      Index     : UINT;     // Byte index. SK: Index bajtu.
      BitIndex  : USINT;    // Bit index. SK: Index bitu.
   END_VAR
   Crc := 16#FFFFFFFF;
   IF Length > 0 THEN
      FOR Index := 0 TO Length - 1 DO
         IF (Index >= 36) AND (Index <= 39) THEN
            Current := 0;
         ELSE
            Current := NhApiReadByte(Buffer := Buffer, Offset := Index);
         END_IF;
         Crc := Crc XOR BYTE_TO_DWORD(Current);
         FOR BitIndex := 0 TO 7 DO
            IF (Crc AND 16#00000001) <> 0 THEN
               Crc := SHR(Crc, 1) XOR 16#EDB88320;
            ELSE
               Crc := SHR(Crc, 1);
            END_IF;
         END_FOR;
      END_FOR;
   END_IF;
   NhApiFrameCrc32 := NOT Crc;
END_FUNCTION

FUNCTION NhApiClearBuffer : BOOL
   // Clears the specified number of buffer bytes. SK: Vynuluje zadany pocet bajtov buffera.
   VAR_INPUT
      Buffer : PTR_TO BYTE; // Buffer to clear. SK: Buffer urceny na vynulovanie.
      Length : UINT;        // Number of bytes. SK: Pocet bajtov.
   END_VAR
   VAR
      Index : UINT;         // Index of the cleared byte. SK: Index nulovaneho bajtu.
   END_VAR
   IF Length > 0 THEN
      FOR Index := 0 TO Length - 1 DO
         NhApiWriteByte(Buffer := Buffer, Offset := Index, Value := 0);
      END_FOR;
   END_IF;
   NhApiClearBuffer := TRUE;
END_FUNCTION

FUNCTION NhApiConfigEqual : BOOL
   // Compares two room configuration records. SK: Porovna dva konfiguracne zaznamy miestnosti.
   VAR_INPUT
      A : NH_ROOM_CONFIG; // First config record. SK: Prvy config zaznam.
      B : NH_ROOM_CONFIG; // Second config record. SK: Druhy config zaznam.
   END_VAR
   NhApiConfigEqual := (A.Used = B.Used) AND (A.RoomId = B.RoomId) AND (A.Name = B.Name) AND
      (A.ProjectName = B.ProjectName) AND (A.IconId = B.IconId) AND (A.SortDefault = B.SortDefault);
END_FUNCTION

FUNCTION NhApiStateEqual : BOOL
   // Compares two dynamic room-state records. SK: Porovna dva dynamicke stavove zaznamy miestnosti.
   VAR_INPUT
      A : NH_ROOM_STATE; // First state record. SK: Prvy state zaznam.
      B : NH_ROOM_STATE; // Second state record. SK: Druhy state zaznam.
   END_VAR
   NhApiStateEqual := (A.RoomId = B.RoomId) AND (A.Temperature = B.Temperature) AND
      (A.Humidity = B.Humidity) AND (A.Presence = B.Presence) AND (A.DayPhase = B.DayPhase) AND
      (A.CategoryMask = B.CategoryMask) AND (A.AlarmLevel = B.AlarmLevel) AND
      (A.Online = B.Online) AND (A.Twilight = B.Twilight);
END_FUNCTION

FUNCTION NhApiFindRoom : UINT
   // Finds a room slot by stable RoomId. SK: Najde room slot podla stabilneho RoomId.
   VAR_INPUT
      RoomId : UDINT; // Stable ID to find. SK: Hladane stabilne ID.
   END_VAR
   VAR
      Index : UINT;  // Scanned room slot. SK: Prehladavany room slot.
   END_VAR
   NhApiFindRoom := 0;
   FOR Index := 1 TO NH_API_MAX_ROOMS DO
      IF NhRoomsConfig[Index].Used AND (NhRoomsConfig[Index].RoomId = RoomId) THEN
         NhApiFindRoom := Index;
         RETURN;
      END_IF;
   END_FOR;
END_FUNCTION

FUNCTION NhApiFindFreeRoom : UINT
   // Finds the first free internal room slot. SK: Najde prvy volny interny room slot.
   VAR
      Index : UINT; // Scanned room slot. SK: Prehladavany room slot.
   END_VAR
   NhApiFindFreeRoom := 0;
   FOR Index := 1 TO NH_API_MAX_ROOMS DO
      IF NOT NhRoomsConfig[Index].Used THEN
         NhApiFindFreeRoom := Index;
         RETURN;
      END_IF;
   END_FOR;
END_FUNCTION

FUNCTION NhApiWriteText64 : BOOL
   // Writes text into a fixed 65-byte wire field. SK: Zapise text do pevneho 65-bajtoveho wire pola.
   VAR_INPUT
      Buffer : PTR_TO BYTE; // Destination wire buffer. SK: Cielovy wire buffer.
      Offset : UINT;        // Offset of length and 64 text bytes. SK: Offset dlzky a 64 bajtov textu.
      Value  : STRING[64];  // UTF-8 bytes stored in PLC STRING. SK: UTF-8 bajty ulozene v PLC STRING.
   END_VAR
   VAR
      Source : PTR_TO BYTE; // First PLC STRING byte. SK: Prvy bajt PLC STRING.
      Index  : USINT;       // Text byte index. SK: Index textoveho bajtu.
      Count  : USINT;       // Actual byte count. SK: Skutocny pocet bajtov.
   END_VAR
   Count := INT_TO_USINT(LEN(Value));
   IF Count > 64 THEN Count := 64; END_IF;
   NhApiWriteByte(Buffer := Buffer, Offset := Offset, Value := USINT_TO_BYTE(Count));
   Source := ADR(Value);
   FOR Index := 0 TO 63 DO
      IF Index < Count THEN
         NhApiWriteByte(Buffer := Buffer, Offset := Offset + 1 + USINT_TO_UINT(Index),
            Value := NhApiReadByte(Buffer := Source, Offset := USINT_TO_UINT(Index)));
      ELSE
         NhApiWriteByte(Buffer := Buffer, Offset := Offset + 1 + USINT_TO_UINT(Index), Value := 0);
      END_IF;
   END_FOR;
   NhApiWriteText64 := TRUE;
END_FUNCTION

FUNCTION NhApiReadText64 : STRING[64]
   // Reads text from a fixed 65-byte wire field. SK: Precita text z pevneho 65-bajtoveho wire pola.
   VAR_INPUT
      Buffer : PTR_TO BYTE; // Source wire buffer. SK: Zdrojovy wire buffer.
      Offset : UINT;        // Offset of length and 64 text bytes. SK: Offset dlzky a 64 bajtov textu.
   END_VAR
   VAR
      Destination : PTR_TO BYTE; // First byte of result PLC STRING. SK: Prvy bajt vysledneho PLC STRING.
      Index       : USINT;       // Text byte index. SK: Index textoveho bajtu.
      Count       : USINT;       // Declared byte count. SK: Deklarovany pocet bajtov.
   END_VAR
   Count := BYTE_TO_USINT(NhApiReadByte(Buffer := Buffer, Offset := Offset));
   IF Count > 64 THEN Count := 64; END_IF;
   Destination := ADR(NhApiReadText64);
   FOR Index := 0 TO 63 DO
      IF Index < Count THEN
         NhApiWriteByte(Buffer := Destination, Offset := USINT_TO_UINT(Index),
            Value := NhApiReadByte(Buffer := Buffer, Offset := Offset + 1 + USINT_TO_UINT(Index)));
      ELSE
         NhApiWriteByte(Buffer := Destination, Offset := USINT_TO_UINT(Index), Value := 0);
      END_IF;
   END_FOR;
END_FUNCTION

FUNCTION NhApiWriteConfigRecord : BOOL
   // Serializes one room configuration record. SK: Serializuje jeden konfiguracny zaznam miestnosti.
   VAR_INPUT
      Buffer : PTR_TO BYTE;      // Destination wire buffer. SK: Cielovy wire buffer.
      Offset : UINT;             // Record start offset. SK: Offset zaciatku zaznamu.
      Record : NH_ROOM_CONFIG;   // Config record to serialize. SK: Config zaznam na serializaciu.
   END_VAR
   NhApiWriteU32(Buffer := Buffer, Offset := Offset, Value := Record.RoomId);
   NhApiWriteU16(Buffer := Buffer, Offset := Offset + 4, Value := Record.IconId);
   NhApiWriteU16(Buffer := Buffer, Offset := Offset + 6, Value := Record.SortDefault);
   NhApiWriteText64(Buffer := Buffer, Offset := Offset + 8, Value := Record.Name);
   NhApiWriteText64(Buffer := Buffer, Offset := Offset + 73, Value := Record.ProjectName);
   NhApiWriteConfigRecord := TRUE;
END_FUNCTION

FUNCTION NhApiReadConfigRecord : BOOL
   // Deserializes one room configuration record. SK: Deserializuje jeden konfiguracny zaznam miestnosti.
   VAR_INPUT
      Buffer : PTR_TO BYTE;      // Source wire buffer. SK: Zdrojovy wire buffer.
      Offset : UINT;             // Record start offset. SK: Offset zaciatku zaznamu.
   END_VAR
   VAR_IN_OUT
      Record : NH_ROOM_CONFIG;   // Decoded config record. SK: Dekodovany config zaznam.
   END_VAR
   Record.Used := TRUE;
   Record.RoomId := NhApiReadU32(Buffer := Buffer, Offset := Offset);
   Record.IconId := NhApiReadU16(Buffer := Buffer, Offset := Offset + 4);
   Record.SortDefault := NhApiReadU16(Buffer := Buffer, Offset := Offset + 6);
   Record.Name := NhApiReadText64(Buffer := Buffer, Offset := Offset + 8);
   Record.ProjectName := NhApiReadText64(Buffer := Buffer, Offset := Offset + 73);
   NhApiReadConfigRecord := TRUE;
END_FUNCTION

FUNCTION NhApiWriteStateRecord : BOOL
   // Serializes one dynamic room-state record. SK: Serializuje jeden dynamicky room-state zaznam.
   VAR_INPUT
      Buffer : PTR_TO BYTE;      // Destination wire buffer. SK: Cielovy wire buffer.
      Offset : UINT;             // Record start offset. SK: Offset zaciatku zaznamu.
      Record : NH_ROOM_STATE;    // State record to serialize. SK: State zaznam na serializaciu.
   END_VAR
   NhApiWriteU32(Buffer := Buffer, Offset := Offset, Value := Record.RoomId);
   NhApiWriteReal(Buffer := Buffer, Offset := Offset + 4, Value := Record.Temperature);
   NhApiWriteReal(Buffer := Buffer, Offset := Offset + 8, Value := Record.Humidity);
   NhApiWriteByte(Buffer := Buffer, Offset := Offset + 12, Value := BOOL_TO_BYTE(Record.Presence));
   NhApiWriteU16(Buffer := Buffer, Offset := Offset + 13, Value := Record.DayPhase);
   NhApiWriteU32(Buffer := Buffer, Offset := Offset + 15, Value := DWORD_TO_UDINT(Record.CategoryMask));
   NhApiWriteByte(Buffer := Buffer, Offset := Offset + 19, Value := USINT_TO_BYTE(Record.AlarmLevel));
   NhApiWriteByte(Buffer := Buffer, Offset := Offset + 20, Value := BOOL_TO_BYTE(Record.Online));
   NhApiWriteByte(Buffer := Buffer, Offset := Offset + 21, Value := BOOL_TO_BYTE(Record.Twilight));
   NhApiWriteStateRecord := TRUE;
END_FUNCTION

FUNCTION NhApiReadStateRecord : BOOL
   // Deserializes one dynamic room-state record. SK: Deserializuje jeden dynamicky room-state zaznam.
   VAR_INPUT
      Buffer : PTR_TO BYTE;      // Source wire buffer. SK: Zdrojovy wire buffer.
      Offset : UINT;             // Record start offset. SK: Offset zaciatku zaznamu.
   END_VAR
   VAR_IN_OUT
      Record : NH_ROOM_STATE;    // Decoded state record. SK: Dekodovany state zaznam.
   END_VAR
   Record.RoomId := NhApiReadU32(Buffer := Buffer, Offset := Offset);
   Record.Temperature := NhApiReadReal(Buffer := Buffer, Offset := Offset + 4);
   Record.Humidity := NhApiReadReal(Buffer := Buffer, Offset := Offset + 8);
   Record.Presence := NhApiReadByte(Buffer := Buffer, Offset := Offset + 12) <> 0;
   Record.DayPhase := NhApiReadU16(Buffer := Buffer, Offset := Offset + 13);
   Record.CategoryMask := UDINT_TO_DWORD(NhApiReadU32(Buffer := Buffer, Offset := Offset + 15));
   Record.AlarmLevel := BYTE_TO_USINT(NhApiReadByte(Buffer := Buffer, Offset := Offset + 19));
   Record.Online := NhApiReadByte(Buffer := Buffer, Offset := Offset + 20) <> 0;
   Record.Twilight := NhApiReadByte(Buffer := Buffer, Offset := Offset + 21) <> 0;
   NhApiReadStateRecord := TRUE;
END_FUNCTION
